Staubli VAL3: setFrameData.pgx

program setFrameData(num x_nIndex)
  local bool l_bResult
  local num l_nResult
begin

  l_bResult=userPageConfirm("确定设定坐标系？(点位会随坐标系改变)")

  if l_bResult
    safeTemp:zZoneItem[x_nIndex].fBase.trsf.x=nFrame[0]
    safeTemp:zZoneItem[x_nIndex].fBase.trsf.y=nFrame[1]
    safeTemp:zZoneItem[x_nIndex].fBase.trsf.z=nFrame[2]
    safeTemp:zZoneItem[x_nIndex].fBase.trsf.rx=nFrame[3]
    safeTemp:zZoneItem[x_nIndex].fBase.trsf.ry=nFrame[4]
    safeTemp:zZoneItem[x_nIndex].fBase.trsf.rz=nFrame[5]
    fFrame.trsf=safeTemp:zZoneItem[x_nIndex].fBase.trsf

    l_nResult=safeTemp:libSave()
    if l_nResult==0
      popUpMsg("设定坐标系完成")
    else
      popUpMsg("设定坐标系失败")
    endIf
  endIf
end
